(* Simple Latching Ladder Diagram *)

PROGRAM main
  VAR
    Start AT %IX0.0 : BOOL; (* Simple Hardware Push Button *)
    Stop AT %IX0.1 : BOOL;
    Output AT %QX0.0 : BOOL;
  END_VAR

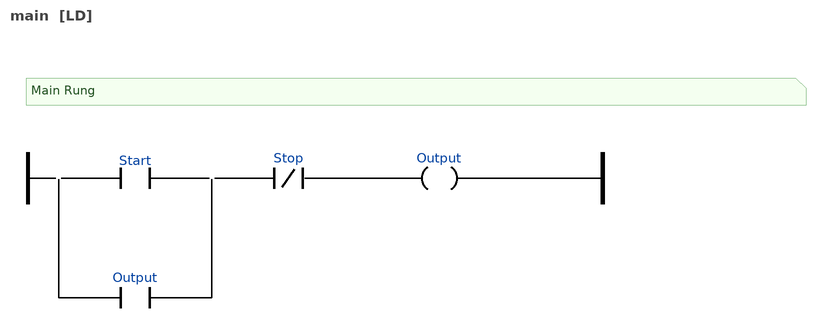
(* LD diagram, written out as Structured Text *)
(* Main Rung *)
Output := (Start OR Output) AND NOT Stop;
END_PROGRAM
